(* EMS UPS 명령 → 세방 UPS 명령 레지스터(0x55) 요청, 온도보상 켜짐 상태 복구 (⑤출력 / 장치: UPS). 2026-11-05.
   기반 없음(신규).
   변경: 없음
   부호·단위: 해당 없음. 명세: C:\gil\UPS\명세서\UPS_명세서.md WR-UPS-01, CF-UPS-03(켜짐 상태). WR-SQ-01은 v2.38에서 폐기
   - 2026-11-12 인터페이스 100.Command: CommandType은 번호 1~26. 번호 n → 세방 맵 명령 주소 99+n (H100~H125)에 0x55
     1 리셋 2 버저 정지 3·4 정류부 ON·OFF 5·6 인버터 ON·OFF 7·8 BBC ON·OFF 9 인버터로 절체 10 바이패스로 절체
     11 부동충전 12 균등충전 13·14 Auto ON·OFF 15 비상 방전 16 주기적 방전 17 펄스 방전 18 방전 취소
     19·20 간헐충전 시작·취소 21·22 온도보상 시작·취소 23·24 ECO 시작·취소 25·26 PRLT 시작·취소
   - 레코드 하나 = 명령 하나. 버전 2의 Delay 대기는 앞에서 FB_EmsCmdGate가 한다
   - 거부: UPS 통신이상이면 모두. UPS 고장(Status b2)이나 e-stop(b3) 중이면 켜기·시작 명령(START_TYPES). 끄기·취소·리셋은 보냄
   - 쓰기 허용(i_bEnable)이 꺼져 있으면 실행하지 않고 Disabled. 장치 명령 1~26, 보고 모드 101 수동·102 자동을 받음
   - 2026-11-17: 드라이버가 바빠 기다리는 동안에도 매 스캔 다시 본다. 고장·e-stop이 생기면 대기 중인 시작 명령을 취소(BadRequest),
     쓰기 허용이 꺼지면 취소(Disabled). 끄기·취소·리셋은 그대로 보낸다
   - Fault 단계 확인은 EMS가 한다 (명세 v2.4). q_bAck는 늘 FALSE
   - 온도보상: 켜 둬야 하는데(iq_stDesired.bTempCompOn) UPS가 꺼져 있으면 i_tRecheck마다 시작 명령을 다시 보낸다.
     i_nMaxFail회 연속으로 켜지지 않으면 q_bEnableMismatch를 켜고 멈춘다. 21·22를 받으면 풀린다 *)
FUNCTION_BLOCK FB_UpsCommand
VAR_INPUT
	i_stCmd			: ST_IfUpsCmd;			// 받은 명령 (번호가 바뀌면 새 명령)
	i_bEnable		: BOOL;					// 장비 쓰기 허용
	i_stUps			: ST_UpsPublish_V1;		// UPS 보고값 (Status b2 고장, b3 e-stop, UPS_ModeStatus b7 온도보상)
	i_bUpsValid		: BOOL;					// UPS 통신 정상
	i_ipUps			: I_Ups;				// 명령 대상
	i_tRequestTimeout : TIME := T#5S;		// 드라이버가 요청을 받지 못하면 실패로 보는 시간
	i_tRecheck		: TIME := T#10S;		// 온도보상 켜짐 상태 확인 주기
	i_nMaxFail		: UINT := 3;			// 켜짐 상태 복구 연속 실패 허용 횟수
END_VAR
VAR_IN_OUT
	iq_stDesired	: ST_UpsDesiredSet;		// 켜짐 상태 보관값 (GVL_PERSIST.g_astUpsDesired[n])
END_VAR
VAR_OUTPUT
	q_bAck				: BOOL;				// Fault 단계 확인. EMS가 하므로 늘 FALSE (v2.4). v2.38부터 MAIN에서 쓰지 않음 (PMS 안 Fault 유지 없앰)
	q_nOperationMode	: UDINT := 1;		// EMS 보고 운전모드: 0 수동(101), 1 자동(102). 시작 기본값 자동
	q_nLastType			: UDINT;			// 마지막으로 받은 명령 번호
	q_eLastResult		: E_UpsResult;		// 마지막 명령 결과
	q_nRejectCount		: UDINT;			// 상태 때문에 거부한 명령 수
	q_nUnknownCount		: UDINT;			// 1~26·101·102 밖의 번호를 받은 수
	q_bDesiredChanged	: BOOL;				// 이 스캔에 켜짐 상태 보관값을 바꿈 (바로 저장 요청)
	q_bEnableMismatch	: BOOL;				// 온도보상 복구 연속 실패 알람
	q_nRestoreCount		: UDINT;			// 온도보상 복구로 시작 명령을 보낸 횟수
END_VAR
VAR
	_nLastSeq		: UDINT;
	_bInit			: BOOL;
	_nPending		: UDINT;				// 드라이버에 넘길 명령 번호 (0 = 없음)
	_tonRequest		: TON;
	_tonRecheck		: TON;
	_nFail			: UINT;
	_bRestoreSent	: BOOL;					// 지난 확인 때 복구 명령을 보냄
	_bFault			: BOOL;
	_bEStop			: BOOL;
	_eCmd			: E_UpsCommand;
	_nNew			: UDINT;
	_bAccepted		: BOOL;
END_VAR
VAR CONSTANT
	MAX_TYPE		: UDINT := 26;		// 번호 1~26 (H100~H125)
	// 고장·e-stop 중 거부하는 켜기·시작 번호: 3 정류부 ON, 5 인버터 ON, 7 BBC ON, 9 인버터로 절체, 11 부동, 12 균등, 13 Auto ON,
	// 15 비상 방전, 16 주기적 방전, 17 펄스 방전, 19 간헐충전, 21 온도보상, 23 ECO, 25 PRLT (비트 n = 번호 n)
	START_TYPES		: DWORD := 16#02ABBAA8;
END_VAR

q_bAck := FALSE;
q_bDesiredChanged := FALSE;
_bFault := i_stUps.Status.2;	// b2 fault
_bEStop := i_stUps.Status.3;	// b3 e-stop

// 처음 스캔: 재시작 전에 받은 명령 번호를 다시 실행하지 않음
IF NOT _bInit THEN
	_bInit := TRUE;
	_nLastSeq := i_stCmd.nSeq;
END_IF

// 1) 새 명령 (1~26 장치, 101 수동·102 자동 보고 모드)
IF i_stCmd.nSeq <> _nLastSeq THEN
	_nLastSeq := i_stCmd.nSeq;
	q_nLastType := i_stCmd.nType;
	_nNew := i_stCmd.nType;
	IF _nNew = 101 OR _nNew = 102 THEN
		// PMS 보고 모드만 변경한다. 세방 Auto ON/OFF(13/14)나 장치 명령은 보내지 않는다.
		IF i_bEnable THEN
			q_nOperationMode := _nNew - 101;
			q_eLastResult := E_UpsResult.Accepted;
		ELSE
			q_eLastResult := E_UpsResult.Disabled;
		END_IF
	ELSIF _nNew = 0 OR _nNew > MAX_TYPE THEN
		q_nUnknownCount := q_nUnknownCount + 1;
		q_eLastResult := E_UpsResult.BadRequest;
	ELSIF NOT i_bUpsValid THEN
		q_nRejectCount := q_nRejectCount + 1;
		q_eLastResult := E_UpsResult.CommUnavailable;
	ELSIF (_bFault OR _bEStop) AND (START_TYPES AND SHL(DWORD#1, UDINT_TO_INT(_nNew))) <> 0 THEN
		q_nRejectCount := q_nRejectCount + 1;	// 고장·e-stop 중 켜기·시작 거부
		q_eLastResult := E_UpsResult.BadRequest;
	ELSIF NOT i_bEnable OR i_ipUps = 0 THEN
		q_eLastResult := E_UpsResult.Disabled;
	ELSE
		_nPending := _nNew;	// 앞의 요청이 남아 있으면 새 명령으로 바꿈 (마지막 명령이 우선)
		q_eLastResult := E_UpsResult.Busy;
	END_IF
END_IF

// 2) 드라이버에 요청. 받아들이면 켜짐 상태 보관값 갱신
_bAccepted := FALSE;
// 2026-11-17: 기다리는 동안 상태가 바뀌면 대기 명령을 취소 (받을 때만 보던 것을 매 스캔 다시 봄)
IF _nPending <> 0 THEN
	IF (_bFault OR _bEStop) AND (START_TYPES AND SHL(DWORD#1, UDINT_TO_INT(_nPending))) <> 0 THEN
		_nPending := 0;
		q_nRejectCount := q_nRejectCount + 1;	// 고장·e-stop이 생겨 시작 명령 취소
		q_eLastResult := E_UpsResult.BadRequest;
	ELSIF NOT i_bEnable OR i_ipUps = 0 THEN
		_nPending := 0;
		q_eLastResult := E_UpsResult.Disabled;
	END_IF
END_IF
_tonRequest(IN := _nPending <> 0, PT := i_tRequestTimeout);
IF _nPending <> 0 THEN
	CASE _nPending OF	// 번호 n → 맵 주소 99+n (E_UpsCommand 값 = 주소)
		1:	_eCmd := E_UpsCommand.Reset;
		2:	_eCmd := E_UpsCommand.BuzzerStop;
		3:	_eCmd := E_UpsCommand.RectifierOn;
		4:	_eCmd := E_UpsCommand.RectifierOff;
		5:	_eCmd := E_UpsCommand.InverterOn;
		6:	_eCmd := E_UpsCommand.InverterOff;
		7:	_eCmd := E_UpsCommand.BbcOn;
		8:	_eCmd := E_UpsCommand.BbcOff;
		9:	_eCmd := E_UpsCommand.ToInverter;
		10:	_eCmd := E_UpsCommand.ToBypass;
		11:	_eCmd := E_UpsCommand.FloatCharge;
		12:	_eCmd := E_UpsCommand.EqualCharge;
		13:	_eCmd := E_UpsCommand.AutoOn;
		14:	_eCmd := E_UpsCommand.AutoOff;
		15:	_eCmd := E_UpsCommand.EmergencyDischarge;
		16:	_eCmd := E_UpsCommand.PeriodicDischarge;
		17:	_eCmd := E_UpsCommand.PulseDischarge;
		18:	_eCmd := E_UpsCommand.CancelDischarge;
		19:	_eCmd := E_UpsCommand.TrickleOn;
		20:	_eCmd := E_UpsCommand.TrickleOff;
		21:	_eCmd := E_UpsCommand.TemperatureOn;
		22:	_eCmd := E_UpsCommand.TemperatureOff;
		23:	_eCmd := E_UpsCommand.EcoOn;
		24:	_eCmd := E_UpsCommand.EcoOff;
		25:	_eCmd := E_UpsCommand.PrltOn;
		26:	_eCmd := E_UpsCommand.PrltOff;
	END_CASE
	IF i_ipUps.M_RequestCommand(_eCmd) THEN
		_bAccepted := TRUE;
		q_eLastResult := E_UpsResult.Accepted;
		CASE _nPending OF
			19:	iq_stDesired.bTrickleOn := TRUE;	q_bDesiredChanged := TRUE;
			20:	iq_stDesired.bTrickleOn := FALSE;	q_bDesiredChanged := TRUE;
			21:	iq_stDesired.bTempCompOn := TRUE;	q_bDesiredChanged := TRUE;	q_bEnableMismatch := FALSE;	_nFail := 0;	_bRestoreSent := FALSE;
			22:	iq_stDesired.bTempCompOn := FALSE;	q_bDesiredChanged := TRUE;	q_bEnableMismatch := FALSE;	_nFail := 0;	_bRestoreSent := FALSE;
		END_CASE
		_nPending := 0;
		_tonRequest(IN := FALSE);
	ELSIF _tonRequest.Q THEN
		_nPending := 0;	// 드라이버가 받지 못함
		q_eLastResult := E_UpsResult.CommUnavailable;
	END_IF
END_IF

// 3) 온도보상 켜짐 상태 복구 (CF-UPS-03)
_tonRecheck(IN := NOT _tonRecheck.Q, PT := i_tRecheck);
IF _tonRecheck.Q AND _nPending = 0 AND NOT _bAccepted THEN
	IF i_stUps.UPS_ModeStatus.7 OR NOT iq_stDesired.bTempCompOn THEN
		_nFail := 0;					// 켜져 있거나 켤 필요 없음
		_bRestoreSent := FALSE;
	ELSIF i_bUpsValid AND i_bEnable AND i_ipUps <> 0 AND NOT _bFault AND NOT _bEStop AND NOT q_bEnableMismatch THEN
		IF _bRestoreSent THEN
			_nFail := _nFail + 1;		// 지난번에 보냈는데 아직 꺼져 있음
		END_IF
		IF _nFail >= i_nMaxFail THEN
			q_bEnableMismatch := TRUE;	// 반복을 멈추고 알람
		ELSIF i_ipUps.M_RequestCommand(E_UpsCommand.TemperatureOn) THEN
			_bRestoreSent := TRUE;
			q_nRestoreCount := q_nRestoreCount + 1;
		END_IF
	END_IF
END_IF

END_FUNCTION_BLOCK

(* stored: Version 1.1.0.1, ProductVersion 3.1.4024.12
   POU FB_UpsCommand: Id {fdd1a924-ca04-4056-888d-a436d42b41d3}, SpecialFunc None *)
